// TIA Portal project "Proyecto_Contador_Rapido_HMI" (V13)

(* hardware
DEVICE "S7-1200 station_1"  S7-1200 Station
   slot 0: "Rack_0"  Rack  V1.0
   slot 1: "PLC_1"  CPU 1214C AC/DC/Rly  6ES7 214-1BE30-0XB0  V2.2
   slot 3: "AQ 1x12BIT_1"  6ES7 232-4HA30-0XB0  V1.0
DEVICE "HMI_1"  KTP600 Basic color PN
   slot 0: "HMI"  HMI  6AV6 647-0AD11-3AX0  11.0.0.0
   slot 1: "HMI_RT_1"  KTP600 Basic color PN  6AV6 647-0AD11-3AX0  11.0.0.0
   slot 5: "HMI_1.IE_CP_1"  Interfaz PROFINET
      slot 1: "Interfaz PROFINET_1"  Interfaz PROFINET
         slot 1: "Port_1"  Port
*)

// ===== PLC "PLC_1"  CPU 1214C AC/DC/Rly =====

VAR_GLOBAL   // PLC tag table "Tabla de variables estándar"
   "Tag_1" AT %ID1000 : DWord;
   "Tag_2" AT %MD200 : DWord;
   "Tag_3" AT %MD300 : DInt;
   "System_Byte" AT %MB1 : Byte;
   "FirstScan" AT %M1.0 : Bool;
   "DiagStatusUpdate" AT %M1.1 : Bool;
   "AlwaysTRUE" AT %M1.2 : Bool;
   "AlwaysFALSE" AT %M1.3 : Bool;
   "Clock_Byte" AT %MB0 : Byte;
   "Clock_5Hz" AT %M0.1 : Bool;
   "Clock_2.5Hz" AT %M0.2 : Bool;
   "Clock_2Hz" AT %M0.3 : Bool;
   "Clock_1.25Hz" AT %M0.4 : Bool;
   "Clock_1Hz" AT %M0.5 : Bool;
   "Clock_0.625Hz" AT %M0.6 : Bool;
   "Clock_0.5Hz" AT %M0.7 : Bool;
   "habilitacion" AT %Q0.0 : Bool;
   "encendido" AT %M10.0 : Bool;
   "parada" AT %M10.1 : Bool;
   "gh" AT %M10.2 : Bool;
   "gah" AT %M10.3 : Bool;
   "velocidad_requerida" AT %MW50 : Int;
   "giro" AT %Q0.1 : Bool;
   "Tag_4" AT %QW80 : Int;
   "Tag_5" AT %MW60 : Word;
   "Tag_6" AT %MD700 : Real;
END_VAR

ORGANIZATION_BLOCK "Main"   // OB1, LAD, ProgramCycle
TITLE = "Main Program Sweep (Cycle)"
{ S7_Optimized_Access := 'FALSE' }
VERSION : 0.1
BEGIN

REGION Network 1
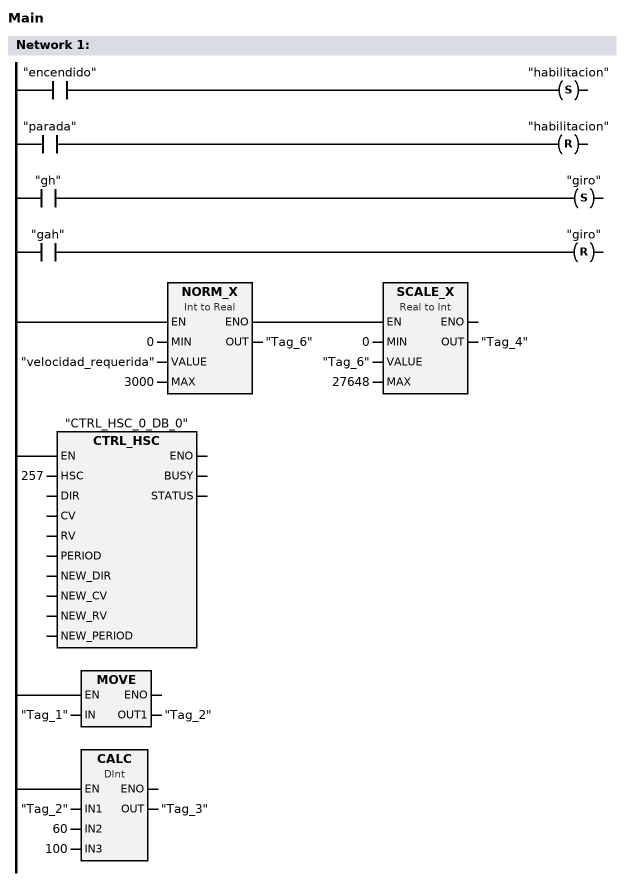
   // ENO of a box is taken as its EN; it also drops when the box reports an error
   IF "encendido" THEN "habilitacion" := TRUE; END_IF;
   IF "parada" THEN "habilitacion" := FALSE; END_IF;
   IF "gh" THEN "giro" := TRUE; END_IF;
   IF "gah" THEN "giro" := FALSE; END_IF;
   "Tag_6" := NORM_X(MIN := 0, VALUE := "velocidad_requerida", MAX := 3000);
   "Tag_4" := SCALE_X(MIN := 0, VALUE := "Tag_6", MAX := 27648);
   "CTRL_HSC_0_DB_0"(HSC := 257);   // CTRL_HSC
   "Tag_2" := "Tag_1";
   CALC(in1 := "Tag_2", in2 := 60, in3 := 100, out => "Tag_3");
END_REGION
END_ORGANIZATION_BLOCK

(* ===== HMI "HMI_RT_1" =====
connection "HMI_Conexión_1": ETHERNET, SMART_S7_1200

HMI tags "Tabla de variables estándar"
   "encendido" : Bool = PLC "encendido", 1 s
   "parada" : Bool = PLC "parada", 1 s
   "velocidad_requerida" : Int = PLC "velocidad_requerida", 1 s
   "Tag_3" : DInt = PLC "Tag_3", 1 s
   "gh" : Bool = PLC "gh", 1 s
   "gah" : Bool = PLC "gah", 1 s

Template "Plantilla_1" 320x240
   Button "Template_Button" at 266,202 size 52x37
   Button "Template_Button_1" at 213,202 size 52x37
   Button "Template_Button_2" at 160,202 size 52x37
   Button "Template_Button_3" at 107,202 size 52x37
   Button "Template_Button_4" at 54,202 size 52x37
   Button "Template_Button_5" at 1,202 size 52x37

screen "Imagen raíz" 320x240, template "Plantilla_1"
   Button "Botón_1" at 15,11 size 96x32
   Button "Botón_2" at 16,61 size 96x32
   IOField "Campo ES_1" at 19,163 size 96x23
   Bar "Barra_1" at 260,67 size 60x120
   Button "Botón_3" at 131,10 size 96x32
   Button "Botón_4" at 128,61 size 96x32
*)